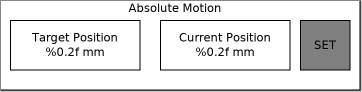
VISUALIZATION ABSOLUTE_MOTION  // 362x92
    Rectangle (-10,0 370x90), "Absolute Motion"
    Rectangle (10,20 130x50), "Target Position %0.2f mm", text variable: MAIN.TargetPosition
        OnMouseDown: write the text variable via VisuDialogs.Numpad, min MAIN.Track.LimitNeg, max MAIN.Track.LimitPos, title 'Input Desired Position'
    Rectangle (160,20 130x50), "Current Position %0.2f mm", text variable: MAIN.Track.CurrentPosition
    Rectangle (300,20 50x50), "SET", colour toggle: MAIN.Track.EnableMotion
        tap MAIN.Track.EnableMotion
END_VISUALIZATION

(* stored: Version 1.1.0.1, ProductVersion 3.1.4024.16
   Visu ABSOLUTE_MOTION: Id {28fd5a54-ddce-46ed-9411-e06e578d2ec3} *)
